(* IEC 61131-3 sources: llm-plc-st-eval/data/processed_definitivo/gpt-4o-2024-08-06/I4/zero_shot, 3 files *)

(* ---- ejec_1.st ---- *)
FUNCTION_BLOCK FB_EstrellaTriangulo
VAR_INPUT
    btnMarcha : BOOL; // Botón de marcha
    btnParo : BOOL;   // Botón de paro
END_VAR

VAR_OUTPUT
    kM : BOOL := FALSE; // Contactor principal
    kY : BOOL := FALSE; // Contactor estrella
    kD : BOOL := FALSE; // Contactor triángulo
END_VAR

VAR
    timerEstrella : TON; // Temporizador para el modo estrella
    timerMuerto : TON;   // Temporizador para el tiempo muerto
    estado : INT := 0;   // Estado del proceso
END_VAR

// Implementación del arranque estrella-triángulo
IF btnParo THEN
    // Si se presiona el botón de paro, desactivar todos los contactores y resetear el estado
    kM := FALSE;
    kY := FALSE;
    kD := FALSE;
    estado := 0;
ELSE
    CASE estado OF
        0: // Estado inicial
            IF btnMarcha THEN
                // Al presionar el botón de marcha, activar el contactor principal y el de estrella
                kM := TRUE;
                kY := TRUE;
                timerEstrella(IN := TRUE, PT := T#8S);
                estado := 1;
            END_IF

        1: // Estado de temporización en estrella
            IF timerEstrella.Q THEN
                // Después de 8 segundos, desactivar el contactor de estrella y activar el temporizador muerto
                kY := FALSE;
                timerEstrella(IN := FALSE);
                timerMuerto(IN := TRUE, PT := T#100MS);
                estado := 2;
            END_IF

        2: // Estado de tiempo muerto
            IF timerMuerto.Q THEN
                // Después de 100 ms, activar el contactor de triángulo
                timerMuerto(IN := FALSE);
                kD := TRUE;
                estado := 3;
            END_IF

        3: // Estado de funcionamiento en triángulo
            // Mantener el estado hasta que se presione el botón de paro
            // No se requiere acción adicional aquí
    END_CASE
END_IF
END_FUNCTION_BLOCK

(* ---- ejec_2.st ---- *)
FUNCTION_BLOCK FB_EstrellaTriangulo
VAR
    // Entradas
    btnMarcha : BOOL;
    btnParo : BOOL;

    // Salidas
    kM : BOOL := FALSE;
    kY : BOOL := FALSE;
    kD : BOOL := FALSE;

    // Variables internas
    estado : INT := 0;
    timerEstrella : TON; // Temporizador para el modo estrella
    timerMuerto : TON;   // Temporizador para el tiempo muerto
END_VAR

// Inicialización de los temporizadores
timerEstrella(IN := FALSE, PT := T#8S);
timerMuerto(IN := FALSE, PT := T#100MS);

// Lógica de control
IF btnParo THEN
    // Si se presiona el botón de paro, desactivar todos los contactores
    kM := FALSE;
    kY := FALSE;
    kD := FALSE;
    estado := 0;
ELSIF btnMarcha THEN
    CASE estado OF
        0: // Estado inicial
            kM := TRUE; // Activar contactor principal
            kY := TRUE; // Activar contactor estrella
            timerEstrella(IN := TRUE); // Iniciar temporizador estrella
            estado := 1;

        1: // Esperando que termine el temporizador estrella
            IF timerEstrella.Q THEN
                kY := FALSE; // Desactivar contactor estrella
                timerEstrella(IN := FALSE); // Reiniciar temporizador estrella
                timerMuerto(IN := TRUE); // Iniciar temporizador muerto
                estado := 2;
            END_IF

        2: // Esperando que termine el tiempo muerto
            IF timerMuerto.Q THEN
                kD := TRUE; // Activar contactor triángulo
                timerMuerto(IN := FALSE); // Reiniciar temporizador muerto
                estado := 3;
            END_IF

        3: // Estado final, contactor triángulo activado
            // Mantener el estado hasta que se presione btnParo
            // o se desactive btnMarcha
            IF NOT btnMarcha THEN
                kM := FALSE;
                kD := FALSE;
                estado := 0;
            END_IF
    END_CASE
ELSE
    // Si btnMarcha no está activo, asegurarse de que todo esté apagado
    kM := FALSE;
    kY := FALSE;
    kD := FALSE;
    estado := 0;
END_IF
END_FUNCTION_BLOCK

(* ---- ejec_3.st ---- *)
FUNCTION_BLOCK FB_EstrellaTriangulo
VAR
    // Entradas
    btnMarcha : BOOL;
    btnParo : BOOL;

    // Salidas
    kM : BOOL := FALSE;
    kY : BOOL := FALSE;
    kD : BOOL := FALSE;

    // Variables internas
    estado : INT := 0;
    timerEstrella : TON; // Temporizador para el modo estrella
    timerMuerto : TON;   // Temporizador para el tiempo muerto
END_VAR

// Configuración de los temporizadores
timerEstrella(IN := FALSE, PT := T#8S);
timerMuerto(IN := FALSE, PT := T#100MS);

// Lógica de control
IF btnParo THEN
    // Si se presiona el botón de paro, desactivar todos los contactores
    kM := FALSE;
    kY := FALSE;
    kD := FALSE;
    estado := 0;
ELSIF btnMarcha THEN
    CASE estado OF
        0: // Estado inicial
            kM := TRUE;
            kY := TRUE;
            timerEstrella(IN := TRUE);
            estado := 1;

        1: // Esperando el tiempo de estrella
            IF timerEstrella.Q THEN
                kY := FALSE;
                timerEstrella(IN := FALSE);
                timerMuerto(IN := TRUE);
                estado := 2;
            END_IF

        2: // Tiempo muerto entre estrella y triángulo
            IF timerMuerto.Q THEN
                kD := TRUE;
                timerMuerto(IN := FALSE);
                estado := 3;
            END_IF

        3: // Modo triángulo
            // Mantenerse en este estado hasta que se presione el botón de paro
            // No se requiere acción adicional
    END_CASE
ELSE
    // Si no se presiona ningún botón, asegurar que los contactores estén desactivados
    kM := FALSE;
    kY := FALSE;
    kD := FALSE;
    estado := 0;
END_IF
END_FUNCTION_BLOCK
